(* IEC 61131-3 sources: guidance-for-physical-ai-production-designer-on-aws/source/plan2cell/crates/bt2plc/templates/codesys/device/GVL, 2 files *)

(* ---- GVL_DeviceParams.st ---- *)
(*
 * GVL_DeviceParams
 * PROFINET device identity parameters.
 * Device simulator {{ROBOT_TAG}} ({{ROBOT_NS}}, station {{STATION}}), cell {{CELL_ID}}. Generated by {{GENERATOR}}.
 *
 * These parameters configure how the CODESYS PROFINET Device presents itself
 * on the network. They MUST match what the Siemens PLC expects (from the GSDML).
 *
 * In CODESYS, these are typically set via:
 *   1. The "PROFINET Device IEC Objects" tab in the device editor
 *   2. Or programmatically by writing to the device parameter structure
 *
 * The CODESYS PROFINET Device stack reads these at startup and uses them
 * in DCP responses and during the PROFINET connection establishment.
 *
 * IMPORTANT: The default CODESYS values (VendorId=0x02CC, DeviceId=0x1017)
 * will NOT work with the Siemens PLC that expects KUKA (0x019B / 0x0301).
 * You MUST override them.
 *)

{attribute 'qualified_only'}
VAR_GLOBAL CONSTANT
    (* === KUKA VKRCnexxt Device Identity === *)
    (* These values come from GSDML-V2.25-KUKA-Roboter-GmbH-VKR C4-Device-V1.0 *)

    VENDOR_ID           : UINT        := 16#019B;                 (* KUKA Roboter GmbH *)
    DEVICE_ID           : UINT        := 16#0301;                 (* VKR C4 Device *)
    STATION_TYPE        : STRING(240) := 'KUKA VKR C4';           (* Station type string *)
    DEVICE_TYPE         : STRING(28)  := 'KUKA VKR C4';           (* Device type string *)
    ORDER_ID            : STRING(20)  := 'KUKA VKRC nexxt';       (* Order number *)
    HW_REVISION         : UINT        := 1;                       (* Hardware revision *)
    SW_REV_PREFIX       : USINT       := 16#56;                   (* 'V' in ASCII *)
    SW_REV_MAJOR        : UINT        := 8;                       (* V8.x *)
    SW_REV_MINOR        : UINT        := 2;                       (* x.2 *)
    SW_REV_PATCH        : UINT        := 0;                       (* x.x.0 *)

    (* === Module Identification Numbers (from GSDML) === *)
    MODULE_IDENT_DAP    : DWORD       := DWORD#16#00000301;       (* DAP - Slot 0 *)
    MODULE_IDENT_FDIO64 : DWORD       := DWORD#16#0000008F;       (* PROFIsafe - Slot 1 *)
    MODULE_IDENT_DIO256 : DWORD       := DWORD#16#00001000;       (* VASS telegram - Slot 2 *)
    SUBMODULE_IDENT     : DWORD       := DWORD#16#00000001;       (* Submodule ident (all slots) *)

    (* === PROFIsafe Parameters (Slot 1) === *)
    (* These must match the F-parameter record in the PLC safety configuration *)
    F_SIL_LEVEL         : UINT        := 3;                       (* SIL 3 *)
    F_CRC_LENGTH        : UINT        := 3;                       (* 3-byte CRC *)
    F_WD_TIME_DEFAULT   : UINT        := 500;                     (* Watchdog 500ms *)
    F_BLOCK_ID          : UINT        := 0;                       (* Block ID *)
    F_PAR_CRC_DEFAULT   : UINT        := 16#FF59;                 (* Default F_Par_CRC = 65369 *)
END_VAR

(* ---- GVL_IO.st ---- *)
(*
 * GVL_IO
 * Global variable list for the PROFINET device I/O mapping.
 * Device simulator {{ROBOT_TAG}} ({{ROBOT_NS}}, station {{STATION}}), cell {{CELL_ID}}. Generated by {{GENERATOR}}.
 *
 * These variables are mapped to the PROFINET device modules via the I/O Mapping tab.
 * Do NOT use AT addresses - the mapping is done in the device configuration.
 * Only PLC_PRG accesses this GVL: it copies the commands into local images and writes
 * the robot status back as a whole array / as scalars (the FBs never touch GVL_IO).
 *
 * Module mapping (set in I/O Mapping tab of each module):
 *   SafeIO_FDIO64 (Slot 1):
 *     "8 safe digital inputs" channels  -> GVL_IO.bySafeIn0..bySafeIn7
 *     "8 safe digital outputs" channels -> GVL_IO.bySafeOut0..bySafeOut7
 *
 *   VASS_DIO256 (Slot 2):
 *     Input channel  -> GVL_IO.aVassInputData
 *     Output channel -> GVL_IO.aVassOutputData
 *)

{attribute 'qualified_only'}
VAR_GLOBAL
    (* ========================================================================
       SLOT 1 - PROFIsafe FDIO64 Module
       8 individual USINT/BYTE channels per direction
       Map each one to the corresponding "8 safe digital inputs/outputs" row
       ======================================================================== *)

    (* Safe Inputs: Robot -> PLC (mapped to "8 safe digital inputs" channels) *)
    bySafeIn0       : BYTE;     (* Safe input byte 0: Drive status *)
    bySafeIn1       : BYTE;     (* Safe input byte 1: Gate/protection *)
    bySafeIn2       : BYTE;     (* Safe input byte 2: STO/SS1/SS2/SOS/SLS *)
    bySafeIn3       : BYTE;     (* Safe input byte 3: User *)
    bySafeIn4       : BYTE;     (* Safe input byte 4: User *)
    bySafeIn5       : BYTE;     (* Safe input byte 5: User *)
    bySafeIn6       : BYTE;     (* Safe input byte 6: User *)
    bySafeIn7       : BYTE;     (* Safe input byte 7: User *)

    (* Safe Outputs: PLC -> Robot (mapped to "8 safe digital outputs" channels) *)
    bySafeOut0      : BYTE;     (* Safe output byte 0: Drive enable, E-Stop, SS1/SS2 *)
    bySafeOut1      : BYTE;     (* Safe output byte 1: Zone enables *)
    bySafeOut2      : BYTE;     (* Safe output byte 2: User *)
    bySafeOut3      : BYTE;     (* Safe output byte 3: User *)
    bySafeOut4      : BYTE;     (* Safe output byte 4: User *)
    bySafeOut5      : BYTE;     (* Safe output byte 5: User *)
    bySafeOut6      : BYTE;     (* Safe output byte 6: User *)
    bySafeOut7      : BYTE;     (* Safe output byte 7: User *)

    (* ========================================================================
       SLOT 2 - DIO256 VASS Telegram
       32 bytes per direction as arrays
       ======================================================================== *)

    (* VASS Inputs: Robot -> PLC (32 bytes) *)
    aVassInputData      : ARRAY[0..31] OF BYTE;

    (* VASS Outputs: PLC -> Robot (32 bytes) *)
    aVassOutputData     : ARRAY[0..31] OF BYTE;
END_VAR
